Fanuc KAREL source: kb00079.KL

-- PROVISIONAL review KL for V1013-1; original PC SHA256 42b8f84ea59b8b2add990d3311a909dab15b133436d631dda4fd595f8f980639
-- Incomplete behavior may be omitted. Consult companion uncertainty JSON. Do not deploy.
PROGRAM KB00079
%NOLOCKGROUP
BEGIN
  -- UNRESOLVED_PC offsets 5-12; opcodes 9D,23
  -- UNRESOLVED_PC offsets 17-24; opcodes 9D,23
  -- UNRESOLVED_PC offsets 29-36; opcodes 9D,23
  -- UNRESOLVED_PC offsets 41-77; opcodes 27,22,22,22,27,9D,31,7E,4A
  -- UNRESOLVED_PC offsets 82-86; opcodes 7F
END KB00079
